(* IEC 61131-3 sources: RepoSTGen/dataset/project_code/轴控/FB103_全局变量1, 10 files *)

(* ---- GVL_Alarm.st ---- *)
VAR_GLOBAL
	(*轴类*)
	HMI_b调模A轴报警 		AT %MX200.0: BOOL;
	HMI_b调模B轴报警 		AT %MX200.1: BOOL;
	HMI_b送面料轴报警 		AT %MX200.2: BOOL;
	HMI_b取面料轴报警 		AT %MX200.3: BOOL;
	HMI_b横移A轴报警 		AT %MX200.4: BOOL;
	HMI_b升降A轴报警 		AT %MX200.5: BOOL;
	HMI_b横移B轴报警 		AT %MX200.6: BOOL;
	HMI_b升降B轴报警 		AT %MX200.7: BOOL;
	HMI_b出盒轴报警 		AT %MX201.0: BOOL;
	HMI_b铲灰板轴报警 		AT %MX201.1: BOOL;
	HMI_b包面纸轴报警 		AT %MX201.2: BOOL;
	HMI_b上包底轴报警 		AT %MX201.3: BOOL;
	HMI_b折边轴报警 		AT %MX201.4: BOOL;

	(*气类*)
	HMI_b取料气缸报警 		AT %MX201.5: BOOL;
	HMI_b纠偏气缸报警 		AT %MX201.6: BOOL;
	HMI_b挡料定位气缸报警 	AT %MX201.7: BOOL;
	HMI_b翻板气缸报警 		AT %MX202.0: BOOL;
	HMI_b侧压紧气缸报警 	AT %MX202.1: BOOL;
	HMI_b左A包底气缸报警 	AT %MX202.2: BOOL;
	HMI_b右B包底气缸报警 	AT %MX202.3: BOOL;
	HMI_b上包底气缸报警 	AT %MX202.4: BOOL;

	HMI_b下包底气缸报警 	AT %MX202.5: BOOL;
	HMI_b出料推盒气缸报警 	AT %MX202.6: BOOL;
	HMI_b包盒口升降气缸报警 AT %MX202.7: BOOL;
	HMI_b包盒口下压气缸报警 AT %MX203.0: BOOL;
	HMI_b翻底板气缸报警 	AT %MX203.1: BOOL;
	HMI_b推底板气缸报警 	AT %MX203.2: BOOL;
	HMI_b模组吸底板气缸报警 AT %MX203.3: BOOL;

	HMI_b包边纠偏上下气缸报警 AT %MX203.4: BOOL;
	HMI_b包边纠偏左右气缸报警 AT %MX203.5: BOOL;
	HMI_b包边压料气缸报警 	AT %MX203.6: BOOL;
	HMI_b折边上托气缸报警 	AT %MX203.7: BOOL;
	HMI_b包边铲边气缸报警	AT %MX204.0: BOOL;

	HMI_b吸底板真空报警 	AT %MX204.1: BOOL;
	HMI_b取面板真空报警 	AT %MX204.2: BOOL;
	HMI_bA模吸底板真空报警  AT %MX204.3: BOOL;
	HMI_bA模吸面板真空报警  AT %MX204.4: BOOL;
	HMI_bB模吸底板真空报警  AT %MX204.5: BOOL;
    HMI_bB模吸面板真空报警  AT %MX204.6: BOOL;

	(*其它类*)
	HMI_b设备未回零启动报警 AT %MX204.7: BOOL;
	HMI_b设备在手动模式启动报警 AT %MX205.0: BOOL;
	HMI_b急停报警 			AT %MX205.1: BOOL;
	HMI_b总气压报警 		AT %MX205.2: BOOL;

	HMI_b折边工位入料光纤检测异常报警 AT %MX205.3: BOOL;
	HMI_b取料工位入料光纤检测异常报警 AT %MX205.4: BOOL;

END_VAR

(* ---- GVL_AxisVirtual.st ---- *)
VAR_GLOBAL
	FB_AxisControl_AxisVirtual: FB_轴控块;

//轴触发类
	bAxisVirtual_CommunicationOK: BOOL;
	bAxisVirtual_JogFor: BOOL;
	bAxisVirtual_JogBack: BOOL;
	bAxisVirtual_InchForExcute: BOOL;
	bAxisVirtual_InchBackExcute: BOOL;
	bAxisVirtual_StopExcute: BOOL;
	bAxisVirtual_ResetExcute: BOOL;
	bAxisVirtual_AbsExcute: BOOL;
	bAxisVirtual_RelExcute: BOOL;
	bAxisVirtual_VelExcute: BOOL;
	bAxisVirtual_LimitEnable: BOOL;

//轴状态类
	bAxisVirtual_EnableOK: BOOL;
	bAxisVirtual_StopDone: BOOL;
	bAxisVirtual_AbsDone: BOOL;
	bAxisVirtual_RelDone: BOOL;
	bAxisVirtual_VelBusy: BOOL;
	bAxisVirtual_InchBusy: BOOL;
	bAxisVirtual_JogBusy: BOOL;
	bAxisVirtual_AbsBusy: BOOL;
	bAxisVirtual_RelBusy: BOOL;
	bAxisVirtual_Error: BOOL;
	bAxisVirtual_Accing: BOOL;
	bAxisVirtual_Decing: BOOL;
    bAxisVirtual_Standstill: BOOL;

//数据给定类
	rAxisVirtual_JogVelSet: LREAL;
	rAxisVirtual_AbsVelSet: LREAL;
	rAxisVirtual_RelVelSet: LREAL;
	rAxisVirtual_VelVelSet: LREAL;
	rAxisVirtual_InchVelSet: LREAL;

	rAxisVirtual_AbsPositionSet: LREAL;
	rAxisVirtual_RelPositionSet: LREAL;
	rAxisVirtual_InchPositionSet: LREAL;

//数据读取类
    rAxisVirtual_Actposition: LREAL;
	rAxisVirtual_ActVel: LREAL;
	rAxisVirtual_ActTorque: LREAL;

//其它类
    bAxisVirtual_HomeExcute: BOOL;
    bAxisVirtual_HomeBusy: BOOL;
    bAxisVirtual_HomeDone: BOOL;
END_VAR

//HMI_PLC_BOOL映射
VAR_GLOBAL
	HMI_bAxisVirtual_PowerOff: BOOL;
	HMI_bAxisVirtual_JogForward: BOOL;
    HMI_bAxisVirtual_BackForward: BOOL;
END_VAR

//HMI_PLC_Data映射
VAR_GLOBAL
	HMI_rAxisVirtual_ActPos: REAL;
	HMI_rAxisVirtual_ActVel: REAL;
	HMI_rAxisVirtual_AutoVel: REAL;
	HMI_rAxisVirtual_ManualVel: REAL;

	HMI_rAxisVirtual_Lead: REAL;
	HMI_rAxisVirtual_RatioMember: REAL;
	HMI_rAxisVirtual_RatioDenominator: REAL;

	HMI_rAxisVirtual_HomeFastVel: REAL;
	HMI_rAxisVirtual_HomeSlowVel: REAL;
	HMI_rAxisVirtual_LimitPostive: REAL;
	HMI_rAxisVirtual_LimitNegative: REAL;

	HMI_rAxisVirtual_AbsPos1: REAL;
	HMI_rAxisVirtual_AbsPos2: REAL;
	HMI_rAxisVirtual_AbsPos3: REAL;

	HMI_rAxisVirtual_RelPos1: REAL;
	HMI_rAxisVirtual_RelPos2: REAL;
	HMI_rAxisVirtual_RelPos3: REAL;
END_VAR

(* ---- GVL_ButtonAll.st ---- *)
VAR_GLOBAL
	HMI_b总产量清零 AT %MX150.0: BOOL;
	HMI_b初始化 AT %MX150.1: BOOL;
	HMI_b禁用蜂鸣器 AT %MX150.2: BOOL;
END_VAR

(* ---- GVL_ButtonIO.st ---- *)
VAR_GLOBAL
	HMI_b启动                      AT %MX100.0:BOOL;
	HMI_b停止                      AT %MX100.1:BOOL;
	HMI_b复位                      AT %MX100.2:BOOL;
	HMI_b手动模式0自动模式1        AT %MX100.3:BOOL;

	HMI_b取料气缸 				   AT %MX100.4:BOOL;
	HMI_b纠偏气缸  				   AT %MX100.5:BOOL;
	HMI_b挡料定位气缸 			   AT %MX100.6:BOOL;
	HMI_b翻板气缸	 			   AT %MX100.7:BOOL;
	HMI_b侧压紧气缸  			   AT %MX101.0:BOOL;
	HMI_b左A包底气缸 			   AT %MX101.1:BOOL;
	HMI_b右B包底气缸  			   AT %MX101.2:BOOL;
	HMI_b上包底气缸 			   AT %MX101.3:BOOL;

	HMI_b下包底气缸 			  AT %MX101.4:BOOL;
	HMI_b出料推盒气缸  			  AT %MX101.5:BOOL;
	HMI_b包盒口升降气缸			  AT %MX101.6:BOOL;
    HMI_b包盒口下压气缸  		  AT %MX101.7:BOOL;
    HMI_b翻底板气缸 			  AT %MX102.0:BOOL;
	HMI_b推底板气缸 			  AT %MX102.1:BOOL;
	HMI_b模组吸底板气缸  		  AT %MX102.2:BOOL;

	HMI_b包边纠偏上下气缸  		  AT %MX102.3:BOOL;
	HMI_b包边纠偏左右气缸 	      AT %MX102.4:BOOL;
	HMI_b包边压料气缸		      AT %MX102.6:BOOL;
	HMI_b折边上托气缸		      AT %MX102.7:BOOL;
	HMI_b包边铲边气缸 		      AT %MX103.0:BOOL;

	HMI_b吸底板真空 		      AT %MX103.2:BOOL;
	HMI_b取面板真空 		      AT %MX103.3:BOOL;
	HMI_bA模吸底板真空 			  AT %MX103.4:BOOL;
	HMI_bA模吸面板真空 			  AT %MX103.5:BOOL;
	HMI_bB模吸底板真空 			  AT %MX103.6:BOOL;
	HMI_bB模吸面板真空 			  AT %MX103.7:BOOL;

	HMI_b真空泵 				  AT %MX104.0:BOOL;
	HMI_b出料皮带电机 			  AT %MX104.1:BOOL;

END_VAR

(* ---- GVL_Cliyder.st ---- *)
VAR_GLOBAL
	FB_CylinderDisPos取料气缸 		: FB_气缸操作块;
	FB_CylinderDisPos纠偏气缸 		: FB_气缸操作块;
	FB_CylinderDisPos挡料定位气缸 	: FB_气缸操作块;
	FB_CylinderDisPos翻板气缸 	    : FB_气缸操作块;
	FB_CylinderDisPos侧压紧气缸 	: FB_气缸操作块;
	FB_CylinderDisPos左A包底气缸 	: FB_气缸操作块;
	FB_CylinderDisPos右B包底气缸 	: FB_气缸操作块;
	FB_CylinderDisPos上包底气缸 	: FB_气缸操作块;

	FB_CylinderDisPos下包底气缸 	: FB_气缸操作块;
    FB_CylinderDisPos出料推盒气缸 	: FB_气缸操作块;
	FB_CylinderDisPos包盒口升降气缸 : FB_气缸操作块;
	FB_CylinderDisPos包盒口下压气缸 : FB_气缸操作块;
	FB_CylinderDisPos翻底板气缸	    : FB_气缸操作块;
	FB_CylinderDisPos推底板气缸     : FB_气缸操作块;
	FB_CylinderDisPos模组吸底板气缸	: FB_气缸操作块;

	FB_CylinderDisPos包边纠偏上下气缸   : FB_气缸操作块;
	FB_CylinderDisPos包边纠偏左右气缸 	: FB_气缸操作块;
	FB_CylinderDisPos包边压料气缸 	    : FB_气缸操作块;
	FB_CylinderDisPos折边上托气缸 		: FB_气缸操作块;
	FB_CylinderDisPos包边铲边气缸 		: FB_气缸操作块;

END_VAR

(* ---- GVL_Communication.st ---- *)
VAR_GLOBAL

END_VAR

(* ---- GVL_DataAll.st ---- *)
VAR_GLOBAL
	HMI_d设备总产量         AT %MD10251: UDINT;
	HMI_d设备故障码			AT %MD10252: UDINT;
	HMI_d设备运行天数		AT %MD10253: UDINT;
	HMI_d产能				AT %MD10254: UDINT;

	HMI_d设备运行速度       AT %MD15250: REAL;
	HMI_r推底板延时         AT %MD15251: REAL;

	HMI_r盒子长度 			AT %MD15252: REAL;
	HMI_r盒子宽度 			AT %MD15253: REAL;
	HMI_r盒子高度 			AT %MD15254: REAL;
	HMI_r灰板厚度 			AT %MD15255: REAL;
	HMI_r成型间距 			AT %MD15256: REAL;
	HMI_r铲刀原点距离 		AT %MD15257: REAL;
	HMI_r毛刷原点距离 		AT %MD15258: REAL;
END_VAR

(* ---- GVL_DataCylinder.st ---- *)
VAR_GLOBAL
    HMI_r取料气缸打开延时 			AT %MD15500:REAL;
    HMI_r取料气缸关闭延时 			AT %MD15501:REAL;

    HMI_r纠偏气缸打开延时			AT %MD15502:REAL;
    HMI_r纠偏气缸关闭延时 			AT %MD15503:REAL;

    HMI_r挡料定位气缸打开延时 	 	AT %MD15504:REAL;
    HMI_r挡料定位气缸关闭延时 	 	AT %MD15505:REAL;

    HMI_r翻板气缸打开延时 		 	AT %MD15506:REAL;
    HMI_r翻板气缸关闭延时 		 	AT %MD15507:REAL;

    HMI_r侧压紧气缸打开延时 	 	AT %MD15508:REAL;
    HMI_r侧压紧气缸关闭延时 	 	AT %MD15509:REAL;

    HMI_r左A包底气缸打开延时 	 	AT %MD15510:REAL;
    HMI_r左A包底气缸关闭延时 	 	AT %MD15511:REAL;

    HMI_r右B包底气缸打开延时 	 	AT %MD15512:REAL;
    HMI_r右B包底气缸关闭延时 	 	AT %MD15513:REAL;

    HMI_r上包底气缸打开延时   		AT %MD15514:REAL;
    HMI_r上包底气缸关闭延时   		AT %MD15515:REAL;

    HMI_r下包底气缸打开延时   		AT %MD15516:REAL;
    HMI_r下包底气缸关闭延时   		AT %MD15517:REAL;

    HMI_r出料推盒气缸打开延时 	 	AT %MD15518:REAL;
    HMI_r出料推盒气缸关闭延时 	 	AT %MD15519:REAL;

    HMI_r包盒口升降气缸打开延时 	AT %MD15520:REAL;
    HMI_r包盒口升降气缸关闭延时 	AT %MD15521:REAL;

    HMI_r包盒口下压气缸打开延时 	AT %MD15522:REAL;
    HMI_r包盒口下压气缸关闭延时 	AT %MD15523:REAL;

    HMI_r翻底板气缸打开延时 		AT %MD15524:REAL;
    HMI_r翻底板气缸关闭延时 		AT %MD15525:REAL;

    HMI_r推底板气缸打开延时 	 	AT %MD15526:REAL;
    HMI_r推底板气缸关闭延时 	 	AT %MD15527:REAL;

    HMI_r模组吸底板气缸打开延时 	AT %MD15528:REAL;
    HMI_r模组吸底板气缸关闭延时 	AT %MD15529:REAL;

    HMI_r包边纠偏上下气缸打开延时 	AT %MD15530:REAL;
    HMI_r包边纠偏上下气缸关闭延时 	AT %MD15531:REAL;

    HMI_r包边纠偏左右气缸打开延时 	AT %MD15532:REAL;
    HMI_r包边纠偏左右气缸关闭延时 	AT %MD15533:REAL;

    HMI_r包边压料气缸打开延时 	 	AT %MD15534:REAL;
    HMI_r包边压料气缸关闭延时 	 	AT %MD15535:REAL;

    HMI_r折边上托气缸打开延时 	 	AT %MD15536:REAL;
    HMI_r折边上托气缸关闭延时 	 	AT %MD15537:REAL;

    HMI_r包边铲边气缸打开延时 		AT %MD15538:REAL;
    HMI_r包边铲边气缸关闭延时 		AT %MD15539:REAL;

    HMI_r吸底板真空打开延时 	 	AT %MD15540:REAL;
    HMI_r吸底板真空关闭延时 	 	AT %MD15541:REAL;

    HMI_r取面板真空打开延时	     	AT %MD15542:REAL;
    HMI_r取面板真空关闭延时	     	AT %MD15543:REAL;

    HMI_rA模吸底板真空打开延时 	 	AT %MD15544:REAL;
    HMI_rA模吸底板真空关闭延时 	 	AT %MD15545:REAL;

    HMI_rA模吸面板真空打开延时	 	AT %MD15546:REAL;
    HMI_rA模吸面板真空关闭延时	 	AT %MD15547:REAL;

    HMI_rB模吸底板真空打开延时 	 	AT %MD15548:REAL;
    HMI_rB模吸底板真空关闭延时 	 	AT %MD15549:REAL;

    HMI_rB模吸面板真空打开延时	 	AT %MD15550:REAL;
    HMI_rB模吸面板真空关闭延时		AT %MD15551:REAL;

END_VAR

(* ---- GVL_IO.st ---- *)
VAR_GLOBAL

(****************************************************输入****************************************************)
DI_折边工位入料感应 				AT %MX0.0:BOOL;
DI_取料工位入料感应 				AT %MX0.1:BOOL;
DI_手自动选择开关 			        AT %MX0.2:BOOL;
DI_启动按钮 			            AT %MX0.3:BOOL;
DI_停止按钮 	                    AT %MX0.4:BOOL;
DI_复位按钮 					    AT %MX0.5:BOOL;
DI_急停按钮 				        AT %MX0.6:BOOL;

DI_总气压检测			            AT %MX1.0:BOOL;
DI_取面板真空检测 			        AT %MX1.1:BOOL;
DI_吸底板真空检测 			        AT %MX1.2:BOOL;
DI_A吸底板真空检测 					AT %MX1.3:BOOL;
DI_A吸面板真空检测 				    AT %MX1.4:BOOL;
DI_B吸底板真空检测				    AT %MX1.5:BOOL;
DI_B吸面板真空检测 			        AT %MX1.6:BOOL;

DI_取料上下气缸原点 			    AT %MX2.0:BOOL;
DI_取料上下气缸动点 			    AT %MX2.1:BOOL;
DI_入料纠偏气缸原点 			    AT %MX2.2:BOOL;
DI_入料纠偏气缸动点  				AT %MX2.3:BOOL;
DI_翻板气缸原点 				    AT %MX2.4:BOOL;
DI_翻板气缸动点  				    AT %MX2.5:BOOL;
DI_左A包底气缸原点 				    AT %MX2.6:BOOL;
DI_右B包底气缸原点 				    AT %MX2.7:BOOL;

DI_上包底气缸原点			        AT %MX3.0:BOOL;
DI_出料推盒气缸原点 			    AT %MX3.1:BOOL;
DI_出料推盒气缸动点	                AT %MX3.2:BOOL;
DI_包盒口升降气缸原点 		        AT %MX3.3:BOOL;
DI_包盒口升降气缸动点 		        AT %MX3.4:BOOL;
DI_包盒口下压气缸原点 		        AT %MX3.5:BOOL;
DI_包盒口下压气缸动点 			    AT %MX3.6:BOOL;

DI_推底板气缸原点 				    AT %MX4.0:BOOL;
DI_推底板气缸动点 				    AT %MX4.1:BOOL;
DI_翻底板气缸原点 					AT %MX4.2:BOOL;
DI_翻底板气缸动点 				    AT %MX4.3:BOOL;
DI_模组吸底板气缸原点 				AT %MX4.4:BOOL;

DI_调模A步进原点 					AT %MX5.0:BOOL;
DI_调模A步进限位 				    AT %MX5.1:BOOL;
DI_调模B步进原点 				    AT %MX5.2:BOOL;
DI_调模B步进限位 				    AT %MX5.3:BOOL;

(****************************************************输出****************************************************)
(*取料工位*)
DO_取料气缸 					    AT %MX50.0:BOOL;
DO_纠偏气缸 						AT %MX50.1:BOOL;
DO_挡料定位气缸 					AT %MX50.2:BOOL;
(*成型工位*)
DO_翻板气缸							AT %MX50.3:BOOL;
DO_侧压紧气缸 					    AT %MX50.4:BOOL;
DO_左A包底气缸 					    AT %MX50.5:BOOL;
DO_右B包底气缸 					    AT %MX50.6:BOOL;
DO_上包底气缸 						AT %MX50.7:BOOL;

DO_下包底气缸 					    AT %MX51.0:BOOL;
(*出盒工位*)
DO_出料推盒气缸 					AT %MX51.1:BOOL;
DO_包盒口升降气缸					AT %MX51.2:BOOL;
DO_包盒口下压气缸 					AT %MX51.3:BOOL;
(*送底板工位*)
DO_翻底板气缸 						AT %MX51.4:BOOL;
DO_推底板气缸 					    AT %MX51.5:BOOL;
DO_模组吸底板气缸 					AT %MX51.6:BOOL;
(*折边工位*)
DO_包边纠偏上下气缸 				AT %MX52.0:BOOL;
DO_包边纠偏左右气缸 				AT %MX52.1:BOOL;
DO_包边压料气缸 					AT %MX52.2:BOOL;
DO_折边上托气缸 					AT %MX52.3:BOOL;
DO_包边铲边气缸 				    AT %MX52.4:BOOL;

DO_吸底板真空 			            AT %MX53.0:BOOL;
DO_取面板真空 			            AT %MX53.1:BOOL;
DO_A模吸底板真空 				    AT %MX53.2:BOOL;
DO_A模吸面板真空 				    AT %MX53.3:BOOL;
DO_B模吸底板真空 			        AT %MX53.4:BOOL;
DO_B模吸面板真空 			        AT %MX53.5:BOOL;

DO_三色灯红 				        AT %MX54.0:BOOL;
DO_三色灯黄 				        AT %MX54.1:BOOL;
DO_三色灯绿 					    AT %MX54.2:BOOL;
DO_三色灯蜂鸣器					    AT %MX54.3:BOOL;
DO_真空泵 						    AT %MX54.4:BOOL;
DO_出料皮带电机 					AT %MX54.5:BOOL;
DO_升降A轴抱闸释放 					AT %MX54.6:BOOL;
DO_升降B轴抱闸释放					AT %MX54.7:BOOL;

END_VAR

(* ---- GVL_M.st ---- *)
VAR_GLOBAL
	b所有伺服总线通讯OK: BOOL;
	b所有伺服使能OK: BOOL;
	b所有伺服回零OK: BOOL;
	b所有伺服静止中: BOOL;
	b所有气缸原位OK: BOOL;
	b所有气缸关闭OK: BOOL;

	b开机初始化: BOOL;
	b常闭: BOOL := TRUE;
	b常开: BOOL := FALSE;
	b非急停手动模式: BOOL;
	b非急停自动模式: BOOL;

	b开机第一次启动: BOOL;
	b常通: BOOL;

	b自动运行: BOOL;
	b自动互锁: BOOL;
	b设备初始化中: BOOL;
	b轴控初始化: BOOL;
	b设备报警: BOOL;
	b气缸报警: BOOL;
	b真空报警: BOOL;
	b马达报警: BOOL;
	b其它报警: BOOL;

END_VAR
